// TIA Portal V20 export
FUNCTION_BLOCK "01_Alle_Zaehler"   // FB48, FBD
{ S7_Optimized_Access := 'TRUE' }
// stored: MemoryReserve 100, SetENOAutomatically false
   VAR
      Zaehlsignal_Gesamt : Bool;
      Zaehlsignal_IO : Bool;
      Zaehlsignal_NIO : Bool;
      Zaehlsignal_NIO_LabView : Bool;
      "Zaehlsignal_IO_1 Palette 1" : Bool;
      "Zaehlsignal_IO_2 Palette 2" : Bool;
      "Zaehlsignal_IO_3 Palette 3" : Bool;
      "Zaehlsignal_IO_4 Palette 4" : Bool;
      "Zaehlsignal_IO_5 Palette 5" : Bool;
      "Zaehlsignal_NIO_1_Palette NIO" : Bool;
      Zaehlsignal_NIO_2 : Bool;
      Zaehlsignal_NIO_3 : Bool;
      Zaehlsignal_NIO_4 : Bool;
      Zaehlsignal_NIO_5 : Bool;
      Zaehlsignal_NIO_6 : Bool;
   END_VAR
BEGIN

NETWORK
TITLE = Zählerstand Teile Gesamt
      CALL  "Zählerfunktion >1000"
      ( Schichtzaehler_Reset  := "HMI_COM".Reset_Schichtzaehler,
        Auftragszaehler_Reset := "HMI_COM".Reset_Auftragszaehler,
        Schichtzaehler        := "HMI_Statistik"."Zaehler Alle Teile".Schichtzaehler,
        Auftragszaehler       := "HMI_Statistik"."Zaehler Alle Teile".Auftragszaehler,
        Gesamtzaehler         := "HMI_Statistik"."Zaehler Alle Teile".Gesamtzaehler,
        Zaehlsignal           := #Zaehlsignal_Gesamt
      );



NETWORK
TITLE = Zählerstand IO gesamt
      CALL  "Zählerfunktion >1000"
      ( Schichtzaehler_Reset  := "HMI_COM".Reset_Schichtzaehler,
        Auftragszaehler_Reset := "HMI_COM".Reset_Auftragszaehler,
        Schichtzaehler        := "HMI_Statistik"."Zaehler IO Teile".Schichtzaehler,
        Auftragszaehler       := "HMI_Statistik"."Zaehler IO Teile".Auftragszaehler,
        Gesamtzaehler         := "HMI_Statistik"."Zaehler IO Teile".Gesamtzaehler,
        Zaehlsignal           := #Zaehlsignal_IO
      );



NETWORK
TITLE = Zählerstand NIO gesamt

      CALL  "Zählerfunktion >1000"
      ( Schichtzaehler_Reset  := "HMI_COM".Reset_Schichtzaehler,
        Auftragszaehler_Reset := "HMI_COM".Reset_Auftragszaehler,
        Schichtzaehler        := "HMI_Statistik"."Zaehler NIO Teile".Schichtzaehler,
        Auftragszaehler       := "HMI_Statistik"."Zaehler NIO Teile".Auftragszaehler,
        Gesamtzaehler         := "HMI_Statistik"."Zaehler NIO Teile".Gesamtzaehler,
        Zaehlsignal           := #Zaehlsignal_NIO
      );



NETWORK
TITLE = IO Zähler 1

      CALL  "Zählerfunktion >1000"
      ( Schichtzaehler_Reset  := "HMI_COM".Reset_Schichtzaehler,
        Auftragszaehler_Reset := "HMI_COM".Reset_Auftragszaehler,
        Schichtzaehler        := "HMI_Statistik"."IO 1".Schichtzaehler,
        Auftragszaehler       := "HMI_Statistik"."IO 1".Auftragszaehler,
        Gesamtzaehler         := "HMI_Statistik"."IO 1".Gesamtzaehler,
        Zaehlsignal           := #"Zaehlsignal_IO_1 Palette 1"
      );


NETWORK
TITLE = IO Zähler 2

      CALL  "Zählerfunktion >1000"
      ( Schichtzaehler_Reset  := "HMI_COM".Reset_Schichtzaehler,
        Auftragszaehler_Reset := "HMI_COM".Reset_Auftragszaehler,
        Schichtzaehler        := "HMI_Statistik"."IO 2".Schichtzaehler,
        Auftragszaehler       := "HMI_Statistik"."IO 2".Auftragszaehler,
        Gesamtzaehler         := "HMI_Statistik"."IO 2".Gesamtzaehler,
        Zaehlsignal           := #"Zaehlsignal_IO_2 Palette 2"
      );




NETWORK
TITLE = IO Zähler 3

      CALL  "Zählerfunktion >1000"
      ( Schichtzaehler_Reset  := "HMI_COM".Reset_Schichtzaehler,
        Auftragszaehler_Reset := "HMI_COM".Reset_Auftragszaehler,
        Schichtzaehler        := "HMI_Statistik"."IO 3".Schichtzaehler,
        Auftragszaehler       := "HMI_Statistik"."IO 3".Auftragszaehler,
        Gesamtzaehler         := "HMI_Statistik"."IO 3".Gesamtzaehler,
        Zaehlsignal           := #"Zaehlsignal_IO_3 Palette 3"
      );




NETWORK
TITLE = IO Zähler 4

      CALL  "Zählerfunktion >1000"
      ( Schichtzaehler_Reset  := "HMI_COM".Reset_Schichtzaehler,
        Auftragszaehler_Reset := "HMI_COM".Reset_Auftragszaehler,
        Schichtzaehler        := "HMI_Statistik"."IO 4".Schichtzaehler,
        Auftragszaehler       := "HMI_Statistik"."IO 4".Auftragszaehler,
        Gesamtzaehler         := "HMI_Statistik"."IO 4".Gesamtzaehler,
        Zaehlsignal           := #"Zaehlsignal_IO_4 Palette 4"
      );




NETWORK
TITLE = IO Zähler 5

      CALL  "Zählerfunktion >1000"
      ( Schichtzaehler_Reset  := "HMI_COM".Reset_Schichtzaehler,
        Auftragszaehler_Reset := "HMI_COM".Reset_Auftragszaehler,
        Schichtzaehler        := "HMI_Statistik"."IO 5".Schichtzaehler,
        Auftragszaehler       := "HMI_Statistik"."IO 5".Auftragszaehler,
        Gesamtzaehler         := "HMI_Statistik"."IO 5".Gesamtzaehler,
        Zaehlsignal           := #"Zaehlsignal_IO_5 Palette 5"
      );




NETWORK
TITLE = NIO Zähler 1

      CALL  "Zählerfunktion >1000"
      ( Schichtzaehler_Reset  := "HMI_COM".Reset_Schichtzaehler,
        Auftragszaehler_Reset := "HMI_COM".Reset_Auftragszaehler,
        Schichtzaehler        := "HMI_Statistik"."NIO 1".Schichtzaehler,
        Auftragszaehler       := "HMI_Statistik"."NIO 1".Auftragszaehler,
        Gesamtzaehler         := "HMI_Statistik"."NIO 1".Gesamtzaehler,
        Zaehlsignal           := #"Zaehlsignal_NIO_1_Palette NIO"
      );


NETWORK
TITLE = NIO Zähler 2

      CALL  "Zählerfunktion >1000"
      ( Schichtzaehler_Reset  := "HMI_COM".Reset_Schichtzaehler,
        Auftragszaehler_Reset := "HMI_COM".Reset_Auftragszaehler,
        Schichtzaehler        := "HMI_Statistik"."NIO 2".Schichtzaehler,
        Auftragszaehler       := "HMI_Statistik"."NIO 2".Auftragszaehler,
        Gesamtzaehler         := "HMI_Statistik"."NIO 2".Gesamtzaehler,
        Zaehlsignal           := #Zaehlsignal_NIO_2
      );


NETWORK
TITLE = NIO Zähler 3

      CALL  "Zählerfunktion >1000"
      ( Schichtzaehler_Reset  := "HMI_COM".Reset_Schichtzaehler,
        Auftragszaehler_Reset := "HMI_COM".Reset_Auftragszaehler,
        Schichtzaehler        := "HMI_Statistik"."NIO 3".Schichtzaehler,
        Auftragszaehler       := "HMI_Statistik"."NIO 3".Auftragszaehler,
        Gesamtzaehler         := "HMI_Statistik"."NIO 3".Gesamtzaehler,
        Zaehlsignal           := #Zaehlsignal_NIO_3
      );


NETWORK
TITLE = NIO Zähler 4

      CALL  "Zählerfunktion >1000"
      ( Schichtzaehler_Reset  := "HMI_COM".Reset_Schichtzaehler,
        Auftragszaehler_Reset := "HMI_COM".Reset_Auftragszaehler,
        Schichtzaehler        := "HMI_Statistik"."NIO 4".Schichtzaehler,
        Auftragszaehler       := "HMI_Statistik"."NIO 4".Auftragszaehler,
        Gesamtzaehler         := "HMI_Statistik"."NIO 4".Gesamtzaehler,
        Zaehlsignal           := #Zaehlsignal_NIO_4
      );




NETWORK
TITLE = NIO Zähler 5

      CALL  "Zählerfunktion >1000"
      ( Schichtzaehler_Reset  := "HMI_COM".Reset_Schichtzaehler,
        Auftragszaehler_Reset := "HMI_COM".Reset_Auftragszaehler,
        Schichtzaehler        := "HMI_Statistik"."NIO 5".Schichtzaehler,
        Auftragszaehler       := "HMI_Statistik"."NIO 5".Auftragszaehler,
        Gesamtzaehler         := "HMI_Statistik"."NIO 5".Gesamtzaehler,
        Zaehlsignal           := #Zaehlsignal_NIO_5
      );


REGION Network 14 (SCL): Reset Taster
   IF "HMI_COM".Reset_Schichtzaehler THEN
       "HMI_COM".Reset_Schichtzaehler := false;
   END_IF;

   IF "HMI_COM".Reset_Auftragszaehler THEN
       "HMI_COM".Reset_Auftragszaehler := false;
   END_IF;
END_REGION
END_FUNCTION_BLOCK
